Staubli VAL3: HMI_message.pjx

--- HMI_message.pjx ---
Parameters version=s8.15.3Cs9_BS3337 stackSize=5000 millimeterUnit=true
Program file=bind.pgx
Program file=click_logExport.pgx
Program file=click_logSave.pgx
Program file=click_refresh.pgx
Program file=click_refreshAllMsg.pgx
Program file=click_refreshIOMsg.pgx
Program file=click_refreshRobotMsg.pgx
Program file=click_refreshTrajMsg.pgx
Program file=initMsg.pgx
Program file=main.pgx
Program file=start.pgx
Program file=stop.pgx
Data file=HMI_message.dtx
Library alias=rs path=Disk://source/projectSource/robotStatus/robotStatus.pjx
Library alias=util path=Disk://HMI_cs9/HMI_util/HMI_util.pjx

--- HMI_message.dtx ---
bool bToHome
string sRobotMsg[40]
bool bBack
num nMsgType
string sCurrentMsg

--- main.pgx ---
public program main()
  local bool l_bExit
  local string l_sTColor
  local string l_sEColor
  local num l_nClock
  local string l_sFColor
  local string l_sLstMsg
begin
  do
    if util:sPage!="message"
      util:sPage="message"
      call util:loadingPage()
      call bind()
      userPage(util:sPage)
      nMsgType=0
      call initMsg()
      call rs:getLog(sRobotMsg,nMsgType)
      userPageSet("message","btnAllMsg","style.backgroundColor","#33FF33")
      userPageSet("message","btnRobotMsg","style.backgroundColor","#FFFFFF")
      userPageSet("message","btnTrajMsg","style.backgroundColor","#FFFFFF")
      sCurrentMsg=""
    endIf
    if sCurrentMsg!=l_sLstMsg
      l_sLstMsg=sCurrentMsg
      popUpMsg(l_sLstMsg)
      sCurrentMsg=l_sLstMsg=""
    endIf
    if bBack
      bBack=false
      l_bExit=true
    endIf
    delay(0.2)
  until l_bExit==true
end

--- start.pgx ---
program start()
begin
  call main()
end

--- bind.pgx ---
program bind()
begin
  userPageBindClick("message","btnback",bBack,true)
  userPageBind("message","lst1","options",sRobotMsg,size(sRobotMsg),"r")
end

--- click_logExport.pgx ---
program click_logExport()
  local num l_nResult
  local string l_sDate
begin
  l_sDate=getDate("%m_%d %H_%M_%S")
  call rs:saveLog("USB0://LOG_"+l_sDate+"/log",l_nResult)
  if l_nResult!=0
    call rs:saveLog("SP2_USB0://LOG_"+l_sDate+"/log",l_nResult)
    if l_nResult!=0
      popUpMsg("未识别U盘,导出失败:"+toString("",l_nResult))
      return
    endIf
  endIf
  popUpMsg("导出到U盘成功,文件名:LOG_"+l_sDate)
end

--- click_logSave.pgx ---
program click_logSave()
  local num l_nResult
  local string l_sDate
begin
  //  l_sDate=getDate("%m_%d %H_%M_%S")
  //  call rs:saveLog("./LOG_"+l_sDate,l_nResult)
  call rs:saveLog(""+l_sDate,l_nResult)
  if l_nResult!=0
    popUpMsg("保存失败:"+toString("",l_nResult))
    return
  endIf
  popUpMsg("保存成功")
end

--- click_refresh.pgx ---
program click_refresh()
begin
  call initMsg()
  call rs:getLog(sRobotMsg,nMsgType)
end

--- click_refreshAllMsg.pgx ---
program click_refreshAllMsg()
begin
  nMsgType=0
  call initMsg()
  call rs:getLog(sRobotMsg,nMsgType)
  userPageSet("message","btnAllMsg","style.backgroundColor","#33FF33")
  userPageSet("message","btnRobotMsg","style.backgroundColor","#FFFFFF")
  userPageSet("message","btnTrajMsg","style.backgroundColor","#FFFFFF")
  userPageSet("message","btnIOMsg","style.backgroundColor","#FFFFFF")
end

--- click_refreshIOMsg.pgx ---
program click_refreshIOMsg()
begin
  nMsgType=3
  call initMsg()
  call rs:getLog(sRobotMsg,nMsgType)
  userPageSet("message","btnAllMsg","style.backgroundColor","#FFFFFF")
  userPageSet("message","btnRobotMsg","style.backgroundColor","#FFFFFF")
  userPageSet("message","btnTrajMsg","style.backgroundColor","#FFFFFF")
  userPageSet("message","btnIOMsg","style.backgroundColor","#33FF33")
end

--- click_refreshRobotMsg.pgx ---
program click_refreshRobotMsg()
begin
  nMsgType=1
  call initMsg()
  call rs:getLog(sRobotMsg,nMsgType)
  userPageSet("message","btnAllMsg","style.backgroundColor","#FFFFFF")
  userPageSet("message","btnRobotMsg","style.backgroundColor","#33FF33")
  userPageSet("message","btnTrajMsg","style.backgroundColor","#FFFFFF")
  userPageSet("message","btnIOMsg","style.backgroundColor","#FFFFFF")
end

--- click_refreshTrajMsg.pgx ---
program click_refreshTrajMsg()
begin
  nMsgType=2
  call initMsg()
  call rs:getLog(sRobotMsg,nMsgType)
  userPageSet("message","btnAllMsg","style.backgroundColor","#FFFFFF")
  userPageSet("message","btnRobotMsg","style.backgroundColor","#FFFFFF")
  userPageSet("message","btnTrajMsg","style.backgroundColor","#33FF33")
  userPageSet("message","btnIOMsg","style.backgroundColor","#FFFFFF")
end

--- initMsg.pgx ---
program initMsg()
  local num i
begin
  for i=0 to size(sRobotMsg)-1
    sRobotMsg[i]=""
  endFor
end

--- stop.pgx ---
program stop()
begin
end
